INTERFACE iShutterCmdSource

METHOD Process
VAR_IN_OUT
	CmdEvent : stShutterCmdEvent;
END_VAR
END_METHOD

END_INTERFACE

(* stored: Version 1.1.0.1
   Itf iShutterCmdSource: Id {d0feda71-d4be-4b61-af82-bec6d51289df}
   Method Process: Id {469b2737-1c8c-408e-927f-cfef22293fe5} *)
